// TIA Portal V21 export
// export: Created 2026-11-11T00:48:24.0764198Z, ExportSetting WithDefaults, DisplayName Totally Integrated Automation Portal, DisplayVersion V21 Update 3, DisplayName STEP 7 Professional, DisplayVersion V21 Update 3, DisplayName STEP 7 Safety, DisplayVersion V21, DisplayName Tech WebApplication, DisplayVersion V21, DisplayName WinCC Basic/Comfort/Advanced, DisplayVersion V21 Update 3, DisplayName WinCC Unified, DisplayVersion V21 Update 3
FUNCTION_BLOCK "FB_Scl_sl115"   // FB199, SCL
{ S7_Optimized_Access := 'TRUE' }
VERSION : 0.1
// stored: AutoNumber true, IsIECCheckEnabled false, IsRetainMemResEnabled false, MemoryReserve 100, SetENOAutomatically false, UDAEnableTagReadback false
   VAR_INPUT
      v_in_bit0 : Bool;
      v_in_bit1 : Bool;
      v_in_bit2 : Bool;
      v_in_bit3 : Bool;
      v_in_bit4 : Bool;
      v_in_bit5 : Bool;
      v_in_bit6 : Bool;
      v_in_bit7 : Bool;
      v_in_bit8 : Bool;
      v_in_bit9 : Bool;
      v_in_bit10 : Bool;
      v_in_bit11 : Bool;
      v_in_bit12 : Bool;
      v_in_bit13 : Bool;
      v_in_bit14 : Bool;
      v_in_bit15 : Bool;
      v_cmp_step : Byte;
   END_VAR
   VAR_OUTPUT
      v_out : Bool;
      v_err_code : Word;
   END_VAR
   VAR
      inst { S7_SetPoint := 'True'} : IMC;
   END_VAR
BEGIN
   #inst(IN_BIT0 := #v_in_bit0, IN_BIT1 := #v_in_bit1, IN_BIT2 := #v_in_bit2, IN_BIT3 := #v_in_bit3, IN_BIT4 := #v_in_bit4, IN_BIT5 := #v_in_bit5, IN_BIT6 := #v_in_bit6, IN_BIT7 := #v_in_bit7, IN_BIT8 := #v_in_bit8, IN_BIT9 := #v_in_bit9, IN_BIT10 := #v_in_bit10, IN_BIT11 := #v_in_bit11, IN_BIT12 := #v_in_bit12, IN_BIT13 := #v_in_bit13, IN_BIT14 := #v_in_bit14, IN_BIT15 := #v_in_bit15, CMP_STEP := #v_cmp_step, OUT => #v_out, ERR_CODE => #v_err_code);
END_FUNCTION_BLOCK
